{attribute 'enable_dynamic_creation'}
FUNCTION_BLOCK FB_Status
VAR_OUTPUT
	code: E_StatusCode;
	// optional and only set when status is an error. Owned by the status and released with it.
	message: POINTER TO FB_String;
END_VAR

(*
	Releases this status and clears the caller's pointer to it: call it as p^.delete(pSelf:=p).
	pSelf is cleared before the status is freed, so the caller never keeps a dangling pointer.
	A pointer to any other object is refused and left untouched, and nothing is released.
*)
METHOD delete : BOOL
VAR_IN_OUT
	pSelf: POINTER TO FB_Status;
END_VAR
VAR
	_pThis: POINTER TO FB_Status;
END_VAR
_pThis := THIS;
IF pSelf <> _pThis THEN
	RETURN;
END_IF

pSelf := 0;
__DELETE(_pThis);
delete := TRUE;
END_METHOD

//FB_Exit must be implemented explicitly. If there is an implementation, then the
//method is called before the controller removes the code of the function block instance
//(implicit call). The return value is not evaluated.
METHOD FB_Exit: BOOL
VAR_INPUT
    bInCopyCode: BOOL;  // TRUE: the exit method is called in order to leave the instance which will be copied afterwards (online change).  
END_VAR
THIS^.free();
END_METHOD

//FB_Init is always available implicitly and it is used primarily for initialization.
//The return value is not evaluated. For a specific influence, you can also declare the
//methods explicitly and provide additional code there with the standard initialization
//code. You can evaluate the return value.
METHOD FB_Init: BOOL
VAR_INPUT
    bInitRetains: BOOL; // TRUE: the retain variables are initialized (reset warm / reset cold)
    bInCopyCode: BOOL;  // TRUE: the instance will be copied to the copy code afterward (online change)
	code: E_StatusCode;
	message: POINTER TO FB_String;  // ownership transfers to the status; the creator clears its copy. 0 means none
END_VAR
THIS^.code := code;
THIS^.message := message;
END_METHOD

METHOD free
IF THIS^.message <> 0 THEN THIS^.message^.delete(pSelf:=THIS^.message); END_IF
END_METHOD

END_FUNCTION_BLOCK

(* stored: Version 1.1.0.1
   POU FB_Status: Id {7502d296-8874-4aba-89de-396bbd73f912}, SpecialFunc None
   Method delete: Id {c4fd0a50-f9e8-441c-a9e5-5109c1bd765e}
   Method FB_Exit: Id {3b724251-b82f-4054-a000-6e9b3e0640c5}
   Method FB_Init: Id {68bac66e-f7c1-47f4-8264-194ff59c77ef}
   Method free: Id {e7fec7ec-ce4b-48e8-b324-a216f3da6d96} *)
